{attribute 'qualified_only'}
{attribute 'strict'}
TYPE E_LightTower_Type :
(
	eSingleLayer := 0,
	eMultiLayer
);
END_TYPE

(* stored: Version 1.1.0.1, ProductVersion 3.1.4024.15
   DUT E_LightTower_Type: Id {4f70e71b-b390-4168-bb3b-a804dc2d11ad} *)
